FUNCTION_BLOCK RAMP_GENERATOR (* Migrated from IEC 61131-3 ST *)
  (* Standard: 61499-2 *)
  (* Version 1.0, 2026-11-06, st2fb *)
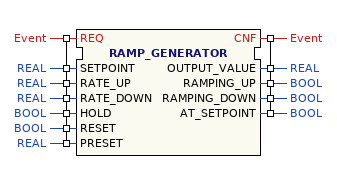
  EVENT_INPUT
    REQ WITH SETPOINT, RATE_UP, RATE_DOWN, HOLD, RESET, PRESET;
  END_EVENT
  EVENT_OUTPUT
    CNF WITH OUTPUT_VALUE, RAMPING_UP, RAMPING_DOWN, AT_SETPOINT;
  END_EVENT
  VAR_INPUT
    SETPOINT : REAL;
    RATE_UP : REAL;
    RATE_DOWN : REAL;
    HOLD : BOOL;
    RESET : BOOL;
    PRESET : REAL;
  END_VAR
  VAR_OUTPUT
    OUTPUT_VALUE : REAL;
    RAMPING_UP : BOOL;
    RAMPING_DOWN : BOOL;
    AT_SETPOINT : BOOL;
  END_VAR
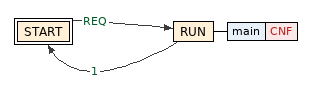
  EC_STATES
    START;
    RUN : main -> CNF;
  END_STATES
  EC_TRANSITIONS
    START TO RUN := REQ;
    RUN TO START := 1;
  END_TRANSITIONS
  ALGORITHM main IN ST:
RAMPING_UP := FALSE;
RAMPING_DOWN := FALSE;
IF RESET THEN
  OUTPUT_VALUE := PRESET;
ELSIF NOT HOLD THEN
  IF OUTPUT_VALUE < SETPOINT THEN
    OUTPUT_VALUE := OUTPUT_VALUE + RATE_UP;
    RAMPING_UP := TRUE;
    IF OUTPUT_VALUE > SETPOINT THEN
      OUTPUT_VALUE := SETPOINT;
    END_IF;
  ELSIF OUTPUT_VALUE > SETPOINT THEN
    OUTPUT_VALUE := OUTPUT_VALUE - RATE_DOWN;
    RAMPING_DOWN := TRUE;
    IF OUTPUT_VALUE < SETPOINT THEN
      OUTPUT_VALUE := SETPOINT;
    END_IF;
  END_IF;
END_IF;
AT_SETPOINT := OUTPUT_VALUE = SETPOINT;
  END_ALGORITHM
END_FUNCTION_BLOCK
